Fanuc KAREL source: kd00011.KL

-- PROVISIONAL review KL for V1013-1; original PC SHA256 bdb5ea416af7bd012bf25451f361af8643e52bef58840e30cfc5118ff287b306
-- Incomplete behavior may be omitted. Consult companion uncertainty JSON. Do not deploy.
PROGRAM KD00011
%NOLOCKGROUP
VAR
  I : INTEGER
  J : INTEGER
  B : BOOLEAN
  R : REAL
  S : STRING[80]
BEGIN
  -- UNRESOLVED_PC offsets 5-6; opcodes 15
  -- UNRESOLVED_PC offsets 11-15; opcodes 7F
END KD00011
